Fanuc KAREL source: kt00534.KL

-- PROVISIONAL review KL for V1013-1; original PC SHA256 0fbf171723c893cc66ae8a9095e5fbd5110149ec77b1773b9e0e8c3b149a9b39
-- Incomplete behavior may be omitted. Consult companion uncertainty JSON. Do not deploy.
PROGRAM KT00534
%NOLOCKGROUP
-- UNRESOLVED_DECL P1 type=000199
-- UNRESOLVED_DECL P2 type=000101
-- UNRESOLVED_DECL OUT type=000101
BEGIN
  -- UNRESOLVED_PC offsets 5-34; opcodes 49,7E,49,60,4A
  -- UNRESOLVED_PC offsets 39-43; opcodes 7F
END KT00534
